// TIA Portal V20 export
// export: Created 2026-10-20T18:55:56.3819718Z, ExportSetting None, DisplayName Totally Integrated Automation Portal, DisplayVersion V20 Update 6, DisplayName TIA Portal Openness, DisplayVersion V20 Update 6, DisplayName TIA Portal Version Control Interface, DisplayVersion V20 Update 6, DisplayName SINAMICS Startdrive Advanced, DisplayVersion V20 SP1, DisplayName SINAMICS Startdrive G130, G150, S120, S150, SINAMICS MV, G220, S200, S210, DisplayVersion V20 SP1, DisplayName SINAMICS Startdrive G110M, G120, G120C, G120D, G120P, G115D, DisplayVersion V20 SP1, DisplayName STEP 7 Professional, DisplayVersion V20 Update 6, DisplayName STEP 7 Safety, DisplayVersion V20 Update 2, DisplayName WinCC Basic/Comfort/Advanced, DisplayVersion V20 Update 6, DisplayName WinCC Unified, DisplayVersion V20 Update 6
VAR_GLOBAL   // PLC tag table "Lock_9"
   Lock_9_Estop_CH1 AT %I1822.2 : Bool;
   Lamps_9 AT %QB1497 : Byte;
   "Solenoid Enable_9" AT %Q1498.0 : Bool;
   Lock_9_Estop_CH2 AT %I1822.3 : Bool;
   Switches_9 AT %IB1496 : Byte;
   Lock_9_Closed_CH2 AT %I1822.1 : Bool;
   "Lock Reset_9" AT %Q1499.0 : Bool;
   Lock_9_Closed_CH1 AT %I1822.0 : Bool;
   Lock_9_Reset_Input3 AT %Q1823.2 : Bool;
   Lock_9_Reset_Input4 AT %Q1823.3 : Bool;
   Lock_9_Reset_Input1 AT %Q1823.0 : Bool;
   Lock_9_Reset_Input2 AT %Q1823.1 : Bool;
   "Lock Position_9" AT %I1572.0 : Bool;
   "Guard Position_9" AT %I1497.0 : Bool;
END_VAR
